FUNCTION_BLOCK "FB_Seq"
VERSION : 0.1
   VAR
      Step : Int;
   END_VAR
BEGIN
	IF #Step = 0 THEN
	    GOTO Done; // PLCA-P006
	END_IF;
	#Step := #Step + 1;
	Done:
	#Step := 3;
END_FUNCTION_BLOCK
